(* IEC 61131-3 sources: 2026_Projet_YGO_ExcavatriceDragage/ARCHIVES/Code/PLC_TESTS/TYPES/ENUMS, 8 files *)

(* ---- E_TestCheckKind.st ---- *)
// ═══════════════════════════════════════════════════════════════
// 🧪 E_TestCheckKind — Enumération des types de checks
// ═══════════════════════════════════════════════════════════════

TYPE E_TestCheckKind :
(
    BOOL_EQUAL     := 0,   // ProbeBool[i] = ExpectedBool
    BOOL_RISING    := 1,   // Front montant de ProbeBool[i]
    BOOL_FALLING   := 2,   // Front descendant de ProbeBool[i]
    DINT_EQUAL     := 3,   // ProbeDint[i] = ExpectedDint
    DINT_NOT_EQUAL := 4,   // ProbeDint[i] <> ExpectedDint
    DINT_IN_RANGE  := 5,   // ExpectedMin <= ProbeDint[i] <= ExpectedMax
    WORD_MASK_ALL  := 6,   // (DINT_TO_WORD(ProbeDint[i]) AND Mask) = Mask
    WORD_MASK_ANY  := 7,   // (DINT_TO_WORD(ProbeDint[i]) AND Mask) <> 0
    WORD_MASK_NONE := 8,   // (DINT_TO_WORD(ProbeDint[i]) AND Mask) = 0
    REAL_IN_RANGE  := 9    // RealMin <= ProbeReal[i] <= RealMax
);
END_TYPE

(* ---- E_TestCheckMode.st ---- *)
// ═══════════════════════════════════════════════════════════════
// 🧪 E_TestCheckMode — Mode d'évaluation des checks
// ═══════════════════════════════════════════════════════════════

TYPE E_TestCheckMode :
(
    CHECK_INSTANT      := 0,  // Vérité exigée au 1er cycle d'évaluation de l'étape (fail sinon)
    CHECK_WAIT_UNTIL   := 1,  // Attendre que ça devienne vrai, tenu StablePT en continu (T#0s = immédiat), borné par TimeoutPT d'étape
    CHECK_INVARIANT    := 2,  // Doit rester vrai CHAQUE cycle de la fenêtre — fail immédiat à la 1re violation
    CHECK_NEVER_DURING := 3   // Ne doit JAMAIS devenir vrai — pass à l'expiration du TimeoutPT d'étape (= la fenêtre)
);
END_TYPE

(* ---- E_TestEventSeverity.st ---- *)
// 🧪 Gravité d'un événement du banc de test
TYPE E_TestEventSeverity :
(
    TEST_EVENT_INFO    := 0,
    TEST_EVENT_WARNING := 1,
    TEST_EVENT_ERROR   := 2
);
END_TYPE

(* ---- E_TestFailAction.st ---- *)
// ═══════════════════════════════════════════════════════════════
// 🧪 E_TestFailAction — Actions à mener en cas d'échec
// ═══════════════════════════════════════════════════════════════

TYPE E_TestFailAction :
(
    FAIL_CONTINUE    := 0,  // Marque l'échec, branche NextOnFail (teardown -> case suivant)
    FAIL_ABORT_SUITE := 1   // Non-récupérable : teardown puis fin de suite
);
END_TYPE

(* ---- E_TestFailReason.st ---- *)
// ═══════════════════════════════════════════════════════════════
// 🧪 E_TestFailReason — Raisons d'échec du test
// ═══════════════════════════════════════════════════════════════

TYPE E_TestFailReason :
(
    FAIL_NONE           := 0,
    FAIL_TIMEOUT        := 1,  // TimeoutPT écoulé sans pass (couvre "trop tard")
    FAIL_CHECK          := 2,  // CHECK_INSTANT faux, ou NEVER_DURING violé
    FAIL_INVARIANT      := 3,  // Invariant multi-étapes violé (voir FailedInvariantId)
    FAIL_WINDOW_EARLY   := 4,  // Pass survenu AVANT MinPT (réaction trop rapide = anormale)
    FAIL_ABORTED        := 5   // Abort commandé ou gate simulation perdu
);
END_TYPE

(* ---- E_TestRunState.st ---- *)
// ═══════════════════════════════════════════════════════════════
// 🧪 E_TestRunState — États d'exécution d'un test
// ═══════════════════════════════════════════════════════════════

TYPE E_TestRunState :
(
    TESTRUN_IDLE    := 0,
    TESTRUN_RUNNING := 1,
    TESTRUN_PASSED  := 2,
    TESTRUN_FAILED  := 3,
    TESTRUN_ABORTED := 4
);
END_TYPE

(* ---- E_TestStimKind.st ---- *)
// ═══════════════════════════════════════════════════════════════
// 🧪 E_TestStimKind — Profils de stimulus instrumentés
// ═══════════════════════════════════════════════════════════════

TYPE E_TestStimKind :
(
    STIM_PULSE_BOOL    := 0,  // Impulsion calibrée PulsePT puis retour auto
    STIM_RAMP_REAL     := 1,  // Rampe linéaire StartReal->TargetReal en RampPT
    STIM_SEQUENCE_REAL := 2   // Profil de valeurs, chacune tenue SeqDwellPT
);
END_TYPE

(* ---- E_TestTerminalState.st ---- *)
// 🧪 État terminal explicite d'une suite ou du séquenceur
TYPE E_TestTerminalState :
(
    TEST_TERMINAL_NONE                 := 0,
    TEST_TERMINAL_DONE                 := 1,
    TEST_TERMINAL_FAILED               := 2,
    TEST_TERMINAL_ABORTED              := 3,
    TEST_TERMINAL_CONFIG_ERROR         := 4,
    TEST_TERMINAL_WATCHDOG_TIMEOUT      := 5,
    TEST_TERMINAL_PRECONDITION_FAILED  := 6  // 🆕 Refus de gate explicite (audit v1.0 C3) — jamais silencieux
);
END_TYPE
